{attribute 'qualified_only'}
VAR_GLOBAL
		Device_1_EtherCAT : Device_1_EtherCAT_49C09C66;
		Device_2_EtherCAT : Device_2_EtherCAT_22CD061B;
		Device_3_EtherCAT : Device_3_EtherCAT_368E547E;
//		Device_4_EtherCAT : Device_4_EtherCAT_07442C6B;
//		Device_5_EtherCAT : Device_5_EtherCAT_0A694E3C;
END_VAR

(* stored: Version 1.2.0.0, ProductVersion 3.1.4024.11
   GVL GVL_iXlinker: Id {38ab9d26-52c2-0cd8-26ba-268c8f1801f0} *)
